(* CODESYS project listofstring.library
   DefaultNamespace: KOSTAL.TC3.Components.listOfString
   DocFormat: reStructuredText
   Description: V2019.2.1.0 - Bugfix: Delete zero pointer
      V2019.2.0.0 - now it is possible to add en empty Line.
      2019.5.0.0 - ListOfString High Performance - Add extended class ListOfString_HP with dynamic storage.
      The temporary load on the router's memory is halved.
   Author: Frank Dümpelmann
   Title: KOSTAL.TC3.Components.listOfString
   Version: 2019.5.0.0
   Company: KOSTAL GmbH & Co.KG
   Placeholder: KOSTAL.TC3.Components.listOfString

Project tree, tasks and I/O mapping:
  libraries: KOSTAL.TC3.Core.functionResponse, 2019.1.0.0 (KOSTAL GmbH & Co.KG); KOSTAL.TC3.Core.Settings, 2019.0.1.0 (KOSTAL GmbH & Co.KG); KOSTAL.TC3.Core.System, 2019.0.0.0 (KOSTAL GmbH & Co.KG); Tc2_Standard, 3.3.3.0 (Beckhoff Automation GmbH); Tc2_System, 3.5.3.0 (Beckhoff Automation GmbH); Tc2_Utilities, 3.3.54.0 (Beckhoff Automation GmbH)
  listOfString_255/
    function block FB_ListOfString_255 [ST]: _stackGetSize, addLine, clear, FB_exit, FB_init, line_GET, line_SET, maxLine, numberOfLines_GET, removeLine
    interface I_ListOfString_255: line_GET, maxLine, numberOfLines_GET
    interface I_ListOfString_255_Owner: addLine, clear, line_GET, line_SET, maxLine, numberOfLines_GET, removeLine
  ListOfString_HP/
    0_Core/
      BaseElement/
        data type P_List
        data type ST_List
      function block FB_Core [ST]: _addItem, _findItem, _findItemByIndex, _insertItem, _removeFromBegin, _removeFromEnd, _removeItem, _removeItemByIndex, _nextItem, _previousItem, _clearResult, _setResultFail, _setResultPass, _checkConsistency, _clear, _NumberOfMember, FB_exit, FB_init
      interface I_Core
      interface I_Core_Owner
    1_Base/
      function block FB_Base [ST]: _FIFO_peek, _FIFO_pop, _FIFO_push, _addMember, _findMember, _findMemberByIndex, _insertMember, _removeFromBegin, _removeFromEnd, _removeMember, _removeMemberByIndex, _clear, FB_exit, FB_init
      interface I_Base
      interface I_Base_Owner
    function block FB_ListOfString_HP [ST]: addLine, clear, line_GET, line_SET, maxLine, maxLine_udi, NumberOfLines, numberOfLines_GET, removeLine
    interface I_ListOfString_HP: maxLine_udi, NumberOfLines
    interface I_ListOfString_HP_Owner: maxLine_udi, NumberOfLines
  Project Information/
    function F_GetCompany [ST]
    function F_GetTitle [ST]
    function F_GetVersion [ST]
  Version/
    global variables Global_Version
*)

// ListOfString_HP/0_Core/BaseElement/P_List
//Pointer to an element of List
TYPE P_List : POINTER TO ST_List; END_TYPE

// ListOfString_HP/0_Core/BaseElement/ST_List
{attribute 'enable_dynamic_creation'}
TYPE ST_List :
	STRUCT
			pNext	 		: P_List;				//Pointer to next Item
			Member			: KOSTAL_TC3_Core_Settings.T_MaxString;	//Text content
			pPrevious : P_List;				//Pointer to previous item
	END_STRUCT
END_TYPE

// Version/Global_Version
{attribute 'TcGenerated'}
{attribute 'no-analysis'}
{attribute 'linkalways'}
// This function has been automatically generated from the project information.
VAR_GLOBAL CONSTANT
	{attribute 'const_non_replaced'}
	stLibVersion_KOSTAL_TC3_Components_listOfString : ST_LibVersion := (iMajor := 2019, iMinor := 5, iBuild := 0, iRevision := 0, nFlags := 1, sVersion := '2019.5.0.0');
END_VAR

// listOfString_255/FB_ListOfString_255
{attribute 'obsolete' := 'Use instead FB_ListOfString_HP'} 
(*

:Author: Frank Dümpelmann <f.duempelmann@kostal.com>, Martin Hundt <m.hundt@kostal.com>
:Date: 2018-11-19

Function
========
Keeps a list of string(255) with a variable number of elements

Usage notes
===============
| Call Method addLine to add a string at the end of the list 
| Call Method getLine to read a string from the list
| numberOfLines_GET returns the actual numer of elements in the list
| List indices are 1-based
| Suitable to implement LIFO or FIFO stacks (see example in fileLogger)

Methods and Properties
======================
| See bottom of this document for a detailed description of each method or property
| Methods starting with an underline(_) are internally used and can be ignored by the user

Usage sample:
=============

.. code:: 

	PROGRAM MAIN
	VAR
		_list	: FB_ListOfString_255;
		_i		: UINT;
		_listContent : ARRAY [1..10] OF STRING(255);
		_filled :BOOL;
	END_VAR
	
	IF NOT _filled THEN	//Add lines to the list ONCE
		_list.addLine('Line 1');
		_list.addLine('Line 2');
		_list.addLine('Line 3');
		_list.addLine('Line 4');
		_list.addLine('Line 5');
		_list.addLine('Line 6');
		_list.removeLine(5);	//Delete line no. 5
		_filled := TRUE;
	END_IF
	
	//Retrieve the lines from the list
	FOR _i:=1 TO _list.numberOfLines_GET() DO
		_listContent[_i] := _list.line_GET(_i);
	END_FOR

*)
FUNCTION_BLOCK PUBLIC FB_ListOfString_255 IMPLEMENTS I_ListOfString_255, I_ListOfString_255_Owner
VAR_INPUT
END_VAR
VAR_OUTPUT
END_VAR

VAR
	_pStack			: POINTER TO KOSTAL_TC3_Core_Settings.T_MaxString;
	_pNewStack	: POINTER TO KOSTAL_TC3_Core_Settings.T_MaxString;
	_line				:	KOSTAL_TC3_Core_Settings.T_MaxString;

	_elements	: UINT;
	_sizeLine	: UDINT;

	_maxLine	:	UINT:= 100;
END_VAR

METHOD PROTECTED _stackGetSize :	UDINT
VAR_INPUT
END_VAR

IF _pStack = 0 THEN
	_stackGetSize:= 0;
ELSE
	_stackGetSize:= SIZEOF(_line) * _elements;
END_IF
END_METHOD

(*
Description
===========
| Adds a line to end of the list
| Parameters:
| 	line: STRING(255): Text to add to the list
| Returns false in case line is empty or list is full
*)

METHOD PUBLIC addLine : BOOL
VAR_INPUT
	newLine	: KOSTAL_TC3_Core_Settings.T_MaxString;
END_VAR

VAR
	_newNumberOfElements	: UINT;
END_VAR

addLine:= FALSE;

//IF newLine = '' THEN RETURN;	END_IF
IF _elements >= _maxLine THEN RETURN;	END_IF

_newNumberOfElements	:= _elements + 1;

_pNewStack:= __NEW(STRING(255), _newNumberOfElements);

IF _elements > 0 THEN
	MEMCPY(destAddr:= ADR(_pNewStack[0]), srcAddr:= ADR(_pStack[0]), n:= _stackGetSize());
END_IF

_pNewStack[_newNumberOfElements - 1]:= newLine;

IF (_pStack <> 0) THEN	__DELETE(_pStack);	END_IF
_elements:= _newNumberOfElements;
_pStack:= __NEW(STRING(255), _elements);

MEMCPY(destAddr:= ADR(_pStack[0]), srcAddr:= ADR(_pNewStack[0]), n:= _stackGetSize());
IF (_pNewStack <> 0) THEN __DELETE(_pNewStack); END_IF

addLine:= TRUE;
END_METHOD

(*
Description
===========
| Clears the list's contents
*)
METHOD PUBLIC clear
VAR_INPUT
END_VAR

IF (_pStack <> 0) THEN __DELETE(_pStack); END_IF
IF (_pNewStack <> 0) THEN __DELETE(_pNewStack); END_IF

_elements:= 0;
END_METHOD

(*
Description
===========
| This method is called automatically
| Do not call manually 
*)
METHOD FB_exit : BOOL
VAR_INPUT
	bInCopyCode : BOOL; // if TRUE, the exit method is called for exiting an instance that is copied afterwards (online change).
END_VAR

IF (_pStack <> 0) THEN __DELETE(_pStack);	END_IF
IF (_pNewStack <> 0) THEN __DELETE(_pNewStack);	END_IF

_elements:= 0;
END_METHOD

(*
Description
===========
| This method is called automatically
| Do not call manually 
*)
METHOD FB_init : BOOL
VAR_INPUT
	bInitRetains : BOOL; // if TRUE, the retain variables are initialized (warm start / cold start)
	bInCopyCode : BOOL;  // if TRUE, the instance afterwards gets moved into the copy code (online change)
END_VAR

IF (_pStack <> 0) THEN __DELETE(_pStack);	END_IF
IF (_pNewStack <> 0) THEN __DELETE(_pNewStack);	END_IF

_elements:= 0;
END_METHOD

(*
Description
===========
| Returns the line at the given index
| Parameters:
| 	numberOfLine: index
*)
METHOD PUBLIC line_GET : KOSTAL_TC3_Core_Settings.T_MaxString
VAR_INPUT
	numberOfLine	:	UINT;	//1..numberOfLines_GET()
END_VAR

line_GET:= '';

IF numberOfLine = 0	THEN	RETURN;	END_IF
IF numberOfLine > _elements THEN	RETURN;	END_IF

line_GET	:=	_pStack[numberOfLine - 1];
END_METHOD

(*
Description
===========
| Returns the line at the given index
| Parameters:
| 	numberOfLine: index
*)
METHOD PUBLIC line_SET : BOOL
VAR_INPUT
	line	: KOSTAL_TC3_Core_Settings.T_MaxString;
	numberOfLine	:	UINT;	//1..numberOfLines_GET()
END_VAR

line_SET:= FALSE;

IF numberOfLine = 0	THEN	RETURN;	END_IF
IF numberOfLine > _elements THEN	RETURN;	END_IF

_pStack[numberOfLine - 1]:= line;

line_SET:= TRUE;
END_METHOD

(*
Description
===========
| **Maximum** number of elements in the list. 
| If the list is full, added lines will be ignored
*)
PROPERTY PUBLIC maxLine : UINT
GET

maxLine:= _maxLine;
END_GET
SET

_maxLine:= maxLine;
END_SET
END_PROPERTY

(*
Description
===========
| Returns the **actual** number of elements in the list
*)
METHOD PUBLIC numberOfLines_GET : UINT
VAR_INPUT
END_VAR

numberOfLines_GET:= _elements;
END_METHOD

(*
Description
===========
| Remove the line with the given index
| Elements after the index move up one position
| Parameters:
| 	index: line to remove
*)

METHOD PUBLIC removeLine
VAR_INPUT
	numberOfLine	:	UINT;	//1..numberOfLines_GET()
END_VAR

VAR
	_indexOfLine		: UINT;
END_VAR


IF numberOfLine = 0 THEN	RETURN;	END_IF
IF numberOfLine > _elements THEN	RETURN;	END_IF

_indexOfLine:= numberOfLine - 1;

_pStack[_indexOfLine]	:= '';

_pNewStack	:=	__NEW(STRING(255), (_elements - 1));

//if not first entry
IF _indexOfLine > 0 THEN
	MEMCPY(destAddr:= ADR(_pNewStack[0]), srcAddr:= ADR(_pStack[0]), n:= SIZEOF(_line) * _indexOfLine);
END_IF

//if not last entry
IF _indexOfLine < _elements - 1 THEN
	MEMCPY(destAddr:= ADR(_pNewStack[_indexOfLine]), srcAddr:= ADR(_pStack[numberOfLine]), n:= SIZEOF(_line) * (_elements - numberOfLine));
END_IF


IF (_pStack <> 0) THEN __DELETE(_pStack);	END_IF

_elements:= _elements - 1;
_pStack:= __NEW(STRING(255), _elements);

MEMCPY(destAddr:= ADR(_pStack[0]), srcAddr:= ADR(_pNewStack[0]), n:= _stackGetSize());
IF (_pNewStack <> 0) THEN __DELETE(_pNewStack);	END_IF
END_METHOD

END_FUNCTION_BLOCK

// ListOfString_HP/FB_ListOfString_HP
(*
	List of String
	HP -High Performance
	The temporary load on the router's memory is halved.
*)
FUNCTION_BLOCK PUBLIC FB_ListOfString_HP EXTENDS FB_Base IMPLEMENTS I_ListOfString_HP, I_ListOfString_HP_Owner
VAR
	_maxLine	: UDINT:= UDINT#16#FFFF_FFFF;
END_VAR

(*
Description
===========
| Adds a line to end of the list
| Parameters:
| 	line: STRING(255): Text to add to the list
| Returns false in case line is empty or list is full
*)
METHOD addLine : BOOL
VAR_INPUT
	newLine	: KOSTAL_TC3_Core_Settings.T_MaxString;
END_VAR

VAR
	_fRes: KOSTAL_TC3_Core_functionResponse.FB_functionResponse;
END_VAR

addLine:= SUPER^._addMember(newLine, _fRes) AND _fRes.success;
END_METHOD

(*
Description
===========
| Clears the list's contents
*)
METHOD clear

SUPER^._clear();
END_METHOD

(*
Description
===========
| Returns the line at the given index
| Parameters:
| 	numberOfLine: index
*)
METHOD line_GET : KOSTAL_TC3_Core_Settings.T_MaxString
VAR_INPUT
	(*1..numberOfLines_GET()*)
	numberOfLine	: UINT;
END_VAR

VAR
	_fRes: KOSTAL_TC3_Core_functionResponse.FB_functionResponse;
END_VAR

_findMemberByIndex(NumberOfLine - 1, line_GET, _fRes);
END_METHOD

(*
Description
===========
| Returns the line at the given index
| Parameters:
| 	numberOfLine: index
*)
METHOD line_SET : BOOL
VAR_INPUT
	line	: KOSTAL_TC3_Core_Settings.T_MaxString;
	(*1..numberOfLines_GET()*)
	numberOfLine	: UINT;
END_VAR

VAR
	_item: P_List;
	_fRes: KOSTAL_TC3_Core_functionResponse.FB_functionResponse;
END_VAR

IF NOT SUPER^._findItemByIndex(numberOfLine - 1, _item, _fRes)	THEN RETURN;	END_IF

IF NOT _fRes.success	THEN RETURN;	END_IF

IF _item = 0 THEN RETURN;	END_IF

_item^.Member:= line;

line_SET:= TRUE;
END_METHOD

(*
Description
===========
| **Maximum** number of elements in the list. 
| If the list is full, added lines will be ignored
*)
PROPERTY maxLine : UINT
GET

IF _maxLine	> UDINT#16#0000_FFFF THEN	maxLine:= UINT#16#FFFF;
ELSE																	maxLine:= UDINT_TO_UINT(_maxLine);
END_IF
END_GET
SET

_maxLine:= UINT_TO_UDINT(maxLine);
END_SET
END_PROPERTY

(*
Description
===========
| **Maximum** number of elements in the list. 
| If the list is full, added lines will be ignored
*)
PROPERTY maxLine_udi : UDINT
GET

maxLine_udi:= _maxLine;
END_GET
SET

_maxLine:= maxLine_udi;
END_SET
END_PROPERTY

PROPERTY PUBLIC NumberOfLines : UDINT
GET

NumberOfLines:= SUPER^._Count;
END_GET
END_PROPERTY


(*
Description
===========
| Returns the **actual** number of elements in the list
*)
METHOD numberOfLines_GET : UINT

IF SUPER^._NumberOfMember > UDINT#16#FFFF THEN	numberOfLines_GET:= UINT#16#FFFF;
ELSE																						numberOfLines_GET:= UDINT_TO_UINT(SUPER^._NumberOfMember);
END_IF
END_METHOD

(*
Description
===========
| Remove the line with the given index
| Elements after the index move up one position
| Parameters:
| 	index: line to remove
*)
METHOD removeLine
VAR_INPUT
	(*1..numberOfLines_GET()*)
	numberOfLine	: UINT;
END_VAR

VAR
	_fRes: KOSTAL_TC3_Core_functionResponse.FB_functionResponse;
END_VAR

SUPER^._removeMemberByIndex(numberOfLine - 1, _fRes);
END_METHOD

END_FUNCTION_BLOCK

// ListOfString_HP/1_Base/FB_Base
(*

| =========================================================================
| List of Items from base Interface {KOSTAL_TC3_Core_System.I_Interface} 
| =========================================================================

..code::

	//In addition to the interface, each item contains the pointer to the previous item 
	//as well as the pointer to the next item in the list.

	TYPE ST_List :
		STRUCT
				pNext			: P_List;
				Line			: KOSTAL_TC3_Core_Settings.T_MaxString;	//Text content
				pPrevious : P_List;
		END_STRUCT
	END_TYPE

============= ======================================= ======================
| The List is defined by (p)Begin and (p)End and also the count of Members 
----------------------------------------------------------------------------
============= ======================================= ======================
 **_pBegin**  >>>>>>>>>>>>>>>>>>>>>>>>>>>>>>>>>>>>>>  **_pEnd**                     
 **Item-1**	    Item-2   Item-3   Item-4  Item-5      **Item-n**                   
============= ======================================= ======================



| =========================================================================
| The Member is an Interface as payload and an access pointer to the        
| previous member and the next member                                      
| ---------------------------------------------------------------------------
| Previous Item ---<<<Pointer-Previous-[Item]-Pointer-Next>>>---NextItem---
| =========================================================================

*)
FUNCTION_BLOCK ABSTRACT FB_Base EXTENDS FB_Core IMPLEMENTS I_Base, I_Base_Owner

VAR
END_VAR

//methode return the Member from begin 
METHOD PROTECTED _FIFO_peek : BOOL
VAR_INPUT
	FoundMember	: REFERENCE TO KOSTAL_TC3_Core_Settings.T_MaxString;	//return value
	Result			: REFERENCE TO KOSTAL_TC3_Core_functionResponse.FB_functionResponse;
END_VAR

_clearResult(Result);

IF 		NOT __ISVALIDREF(FoundMember) THEN _setResultFail(Result, 'FoundMember has no valid reference'); 
ELSE	_FIFO_peek:= _findMemberByIndex(0, FoundMember, Result);
END_IF
END_METHOD

//methode return the Member from begin and remove it from List
METHOD PROTECTED _FIFO_pop : BOOL
VAR_INPUT
	FoundMember	: REFERENCE TO KOSTAL_TC3_Core_Settings.T_MaxString;	//return value
	Result			: REFERENCE TO KOSTAL_TC3_Core_functionResponse.FB_functionResponse;
END_VAR


_clearResult(Result);

_FIFO_pop:= _findMemberByIndex(0, FoundMember, Result);

IF _FIFO_pop THEN	_FIFO_pop:= _removeFromBegin(Result);	END_IF
END_METHOD

//push/add the {Member} to begin from List
METHOD PROTECTED _FIFO_push : BOOL
VAR_INPUT
	Member	: KOSTAL_TC3_Core_Settings.T_MaxString;
	Result	: REFERENCE TO KOSTAL_TC3_Core_functionResponse.FB_functionResponse;
END_VAR


_FIFO_push:= _insertItem(UDINT#0, Member, Result);
END_METHOD

(*
	add new Member to end of list
*)
METHOD PROTECTED _addMember : BOOL

VAR_INPUT
	Member		: KOSTAL_TC3_Core_Settings.T_MaxString;
	Result	: REFERENCE TO KOSTAL_TC3_Core_functionResponse.FB_functionResponse;
END_VAR


VAR
	_Member: KOSTAL_TC3_Core_System.I_Interface;
END_VAR

_addMember:= _addItem(Member, Result);
END_METHOD

(*
	Search for the element {Item} in the list and return {FoundItem} if it is found {_findItem = TRUE}
*)
METHOD PROTECTED _findMember : BOOL
VAR_INPUT
	Member			: KOSTAL_TC3_Core_Settings.T_MaxString;
	FoundMember	: REFERENCE TO KOSTAL_TC3_Core_Settings.T_MaxString;	//return value
	Result			: REFERENCE TO KOSTAL_TC3_Core_functionResponse.FB_functionResponse;
END_VAR

VAR
	_Item		: P_List;
END_VAR

_clearResult(Result);

IF NOT __ISVALIDREF(FoundMember)			THEN _setResultFail(Result, 'FoundItem has no valid reference');	RETURN;	END_IF

_findMember:= _findItem(Member, _Item, Result);

IF NOT _findMember		THEN	RETURN;	END_IF
IF _Item = 0 					THEN	RETURN;	END_IF

FoundMember:= _Item^.Member;
END_METHOD

//find a modul by index  
METHOD PROTECTED _findMemberByIndex : BOOL
VAR_INPUT
	Index				: UDINT;	//index of item
	FoundMember	: REFERENCE TO KOSTAL_TC3_Core_Settings.T_MaxString;	//return value
	Result			: REFERENCE TO KOSTAL_TC3_Core_functionResponse.FB_functionResponse;	//result information
END_VAR

VAR
	_FoundItem	: P_List;
END_VAR

IF NOT __ISVALIDREF(FoundMember)	THEN _setResultFail(Result, 'FoundMember has no valid reference');	RETURN;	END_IF

FoundMember:= '';

_findMemberByIndex:= _findItemByIndex(Index,_FoundItem, Result);

IF NOT _findMemberByIndex THEN RETURN;	END_IF
IF _FoundItem = 0 THEN RETURN;	END_IF

FoundMember:= _FoundItem^.Member;

_findMemberByIndex:= TRUE;
END_METHOD

METHOD PROTECTED _insertMember : BOOL
VAR_INPUT
	Index		: UDINT;	//Index a which shall inserted the {Item}
	Member	: KOSTAL_TC3_Core_Settings.T_MaxString;
	Result	: REFERENCE TO KOSTAL_TC3_Core_functionResponse.FB_functionResponse;
END_VAR

VAR
	_Member: KOSTAL_TC3_Core_System.I_Interface;
END_VAR

_insertMember:= _insertItem(Index, Member, Result);
END_METHOD

(*
	remove Item from begin of list
*)
METHOD PROTECTED _removeFromBegin : BOOL
VAR_INPUT
	Result	: REFERENCE TO KOSTAL_TC3_Core_functionResponse.FB_functionResponse;
END_VAR

_removeFromBegin:= THIS^._removeMemberByIndex(0, Result);
END_METHOD

(*
	remove Item from end of list
*)
METHOD PROTECTED _removeFromEnd : BOOL
VAR_INPUT
	Result	: REFERENCE TO KOSTAL_TC3_Core_functionResponse.FB_functionResponse;
END_VAR

_removeFromEnd:= THIS^._removeMemberByIndex(_Count, Result);
END_METHOD

(*
	remove given {Member} from List
*)
METHOD PROTECTED _removeMember : BOOL
VAR_INPUT
	Member	: KOSTAL_TC3_Core_Settings.T_MaxString;
	Result	: REFERENCE TO KOSTAL_TC3_Core_functionResponse.FB_functionResponse;
END_VAR

VAR
	_Item		: P_List;
	_bFound: BOOL;
END_VAR


_bFound:= _findItem(Member, _Item, Result);

IF NOT _bFound THEN RETURN;	END_IF

_removeMember:= _removeItem(_Item, Result);
END_METHOD

(*
	remove given {Index} from List
*)
METHOD PROTECTED _removeMemberByIndex : BOOL
VAR_INPUT
	Index		: UDINT;
	Result	: REFERENCE TO KOSTAL_TC3_Core_functionResponse.FB_functionResponse;
END_VAR

VAR
	_bFound	: BOOL;
	_Member	: KOSTAL_TC3_Core_Settings.T_MaxString;

END_VAR

IF NOT _findMemberByIndex(Index, _Member, Result)	THEN RETURN;	END_IF

_removeMemberByIndex:= _removeMember(_Member, Result);
END_METHOD

(*
	Delete the complete content of the list
*)
METHOD PROTECTED _clear
VAR_INPUT
END_VAR

WHILE THIS^._pBegin <> 0 DO
    THIS^._removeMember(THIS^._pBegin^.Member, 0);  
END_WHILE
END_METHOD

METHOD FB_exit : BOOL
VAR_INPUT
	bInCopyCode : BOOL; // if TRUE, the exit method is called for exiting an instance that is copied afterwards (online change).
END_VAR

_clear();
END_METHOD

METHOD FB_init : BOOL
VAR_INPUT
	bInitRetains : BOOL; // if TRUE, the retain variables are initialized (warm start / cold start)
	bInCopyCode : BOOL;  // if TRUE, the instance afterwards gets moved into the copy code (online change)
END_VAR

_clear();
END_METHOD

END_FUNCTION_BLOCK

// ListOfString_HP/0_Core/FB_Core
(*

| =========================================================================
| List of Items from base Interface {KOSTAL_TC3_Core_System.I_Interface} 
| =========================================================================

..code::

	//In addition to the interface, each item contains the pointer to the previous item 
	//as well as the pointer to the next item in the list.

	TYPE ST_List :
		STRUCT
				pNext			: P_List;
				iMember		: KOSTAL_TC3_Core_System.I_Interface;	
				pPrevious : P_List;
		END_STRUCT
	END_TYPE

============= ======================================= ======================
| The List is defined by (p)Begin and (p)End and also the count of Members 
----------------------------------------------------------------------------
============= ======================================= ======================
 **_pBegin**  >>>>>>>>>>>>>>>>>>>>>>>>>>>>>>>>>>>>>>  **_pEnd**                     
 **Item-1**	    Item-2   Item-3   Item-4  Item-5      **Item-n**                   
============= ======================================= ======================



| =========================================================================
| The Member is an Interface as payload and an access pointer to the        
| previous member and the next member                                      
| ---------------------------------------------------------------------------
| Previous Item ---<<<Pointer-Previous-[Item]-Pointer-Next>>>---NextItem---
| =========================================================================

*)
FUNCTION_BLOCK ABSTRACT FB_Core IMPLEMENTS I_Core, I_Core_Owner

VAR
	_pBegin	: P_List;	//origin of List
  _pEnd		: P_List;	//end of List
	_Count	: UDINT;	//number of registered Member
END_VAR

(*
	add new item to end of list
*)
METHOD PROTECTED _addItem : BOOL

VAR_INPUT
	Member		: KOSTAL_TC3_Core_Settings.T_MaxString;
	Result	: REFERENCE TO KOSTAL_TC3_Core_functionResponse.FB_functionResponse;
END_VAR

VAR
	_pNewItem	: P_List;
END_VAR
_clearResult(Result);

//IF Item = 0 THEN _setResultFail(Result, 'Parameter Item is empty');	RETURN;	END_IF


//create a new Item
_pNewItem:= __NEW(ST_List);

//If creation failed 
IF _pNewItem = 0 THEN _setResultFail(Result, 'New Item cannot create');	RETURN;	END_IF

//If list is empty
IF THIS^._Count = 0 (*THIS^._pEnd = 0*) THEN THIS^._pBegin:= THIS^._pEnd:= _pNewItem; 
ELSE

	//set new item previous item to actual last item (THIS^._pEnd)
	_pNewItem^.pPrevious:= THIS^._pEnd;
	_pNewItem^.pPrevious^.pNext:= _pNewItem;
 
	THIS^._pEnd:= _pNewItem;
END_IF

THIS^._pEnd^.Member:= Member;
THIS^._Count:= THIS^._Count + UDINT#1;

_setResultPass(Result, 'addItem successful');

_addItem:= TRUE;
END_METHOD

(*
	Search for the element {Item} in the list and return {FoundItem} if it is found {_findItem = TRUE}
*)
METHOD PROTECTED _findItem : BOOL
VAR_INPUT
	Member		: KOSTAL_TC3_Core_Settings.T_MaxString;
	FoundItem	: REFERENCE TO P_List;
	Result		: REFERENCE TO KOSTAL_TC3_Core_functionResponse.FB_functionResponse;
END_VAR

VAR
	_Item		: P_List;
END_VAR
_clearResult(Result);

IF NOT __ISVALIDREF(FoundItem)	THEN _setResultFail(Result, 'FoundItem has no valid reference');	RETURN;	END_IF


_Item := THIS^._pBegin;

WHILE _Item <> 0 DO

	IF _Item^.Member = Member THEN

		FoundItem := _Item;

		_findItem:= TRUE;

		_setResultPass(Result, 'Item found');
		
		RETURN;   

	END_IF
	
	_Item := THIS^._nextItem(_Item, 0);

END_WHILE

//FoundItem:= _Item;

_setResultFail(Result, 'Item not found');

_findItem:= FALSE;
END_METHOD

(*
	Search for the element {Item} in the list and return {FoundItem} if it is found {_findItem = TRUE}
*)
METHOD PROTECTED _findItemByIndex : BOOL
VAR_INPUT
	Index			: UDINT;
	FoundItem	: REFERENCE TO P_List;
	Result		: REFERENCE TO KOSTAL_TC3_Core_functionResponse.FB_functionResponse;
END_VAR

VAR
	_Item		: P_List;
	_udi: UDINT;
END_VAR

_findItemByIndex:= FALSE;

_clearResult(Result);

IF _Count = 0										THEN _setResultFail(Result, 'List is empty');											RETURN;	END_IF
IF Index > (_Count - 1)					THEN _setResultFail(Result, 'Parameter Index is out of range');		RETURN;	END_IF
IF NOT __ISVALIDREF(FoundItem)	THEN _setResultFail(Result, 'FoundItem has no valid reference');	RETURN;	END_IF


_Item := THIS^._pBegin;

IF Index > 0 THEN
	FOR _udi:= 0 TO Index - 1 DO
			_Item := THIS^._nextItem(_Item, 0);
	END_FOR
END_IF

FoundItem:= _Item;

IF FoundItem = 0 THEN
	_setResultFail(Result, 'Item not found');
ELSE	
	_setResultPass(Result, 'Item found');
	_findItemByIndex:= TRUE;
END_IF
END_METHOD

METHOD PROTECTED _insertItem : BOOL
VAR_INPUT
	Index		: UDINT;	//Index a which shall inserted the {Item}
	Member	: KOSTAL_TC3_Core_Settings.T_MaxString;
	Result	: REFERENCE TO KOSTAL_TC3_Core_functionResponse.FB_functionResponse;
END_VAR

VAR
	_pNewItem			: P_List;
	_pExitingItem	: P_List;
END_VAR
_clearResult(Result);

//if List is empty add item 
IF (Index = 0) AND (_Count = 0)	THEN _insertItem:= _addItem(Member, Result);	RETURN;	END_IF

//Index is in list not available 
IF Index > (_Count - 1) THEN _setResultFail(Result, 'Index is out of range');	RETURN;	END_IF

//if index is end of list then add item to end of list 
IF (Index = (_Count - 1)) THEN _insertItem:= _addItem(Member, Result);	RETURN;	END_IF

//try to find item where shall inserted
IF NOT _findItemByIndex(Index, _pExitingItem, Result) THEN RETURN;	END_IF
IF _pExitingItem = 0 THEN _setResultFail(Result, 'Item not available');	RETURN;	END_IF


//create a new Item
_pNewItem:= __NEW(ST_List);

//If creation failed 
IF _pNewItem = 0 THEN _setResultFail(Result, 'New Item cannot create');	RETURN;	END_IF

_pNewItem^.Member:= Member;

_pNewItem^.pNext		:= _pExitingItem;							//set the next item from new item to existing founded item
_pNewItem^.pPrevious:= _pExitingItem^.pPrevious;	//set the previous from existing item to the previous of new item

//if a previous exist then
//set the next from previous from existing item to the previous of new item
IF _pNewItem^.pPrevious <> 0 THEN	_pNewItem^.pPrevious^.pNext:= _pNewItem;	END_IF

_pExitingItem^.pPrevious:= _pNewItem;							//set the previous from existing founded item to  new item

//if inserted at the begin of list, set the begin pointer to new Item
IF THIS^._pBegin = _pExitingItem THEN	THIS^._pBegin:= _pNewItem;	END_IF

THIS^._Count:= THIS^._Count + UDINT#1;

_setResultPass(Result, 'insertItem successful');

_insertItem:= TRUE;
END_METHOD

(*
	remove Item from begin of list
*)
METHOD PROTECTED _removeFromBegin : BOOL
VAR_INPUT
	Result	: REFERENCE TO KOSTAL_TC3_Core_functionResponse.FB_functionResponse;
END_VAR

_removeFromBegin:= THIS^._removeItemByIndex(0, Result);
END_METHOD

(*
	remove Item from end of list
*)
METHOD PROTECTED _removeFromEnd : BOOL
VAR_INPUT
	Result	: REFERENCE TO KOSTAL_TC3_Core_functionResponse.FB_functionResponse;
END_VAR

_removeFromEnd:= THIS^._removeItemByIndex(_Count, Result);
END_METHOD

(*
	remove given {Item} from List
*)
METHOD PROTECTED _removeItem : BOOL
VAR_INPUT
	Item		: P_List;
	Result	: REFERENCE TO KOSTAL_TC3_Core_functionResponse.FB_functionResponse;
END_VAR

_clearResult(Result);

IF Item = 0 THEN _setResultFail(Result, 'Parameter Item is empty');	RETURN;	END_IF

//exist a next member
IF Item^.pNext <> 0 THEN
	//set next members previous Item  to my previous Item
	Item^.pNext^.pPrevious := Item^.pPrevious; 
END_IF

//exist a previous member
IF Item^.pPrevious <> 0 THEN
	//set previous members next Item  to my next Item
	Item^.pPrevious^.pNext := Item^.pNext;
END_IF

//Item is the once member
IF Item = THIS^._pBegin AND Item = THIS^._pEnd THEN
	
	THIS^._pBegin := 0;
	THIS^._pEnd := 0;

ELSIF Item = THIS^._pBegin (*AND Item <> THIS^._pEnd*) THEN

	THIS^._pBegin := Item^.pNext;

ELSIF (*Item <> THIS^._pBegin AND*) Item = THIS^._pEnd THEN

	THIS^._pEnd := Item^.pPrevious;

END_IF

__DELETE(Item);

IF  THIS^._Count > UDINT#0 THEN	THIS^._Count := THIS^._Count - UDINT#1;	
ELSE
	_setResultFail(Result, 'removeItem Counter underflow');
	RETURN;
END_IF

_setResultPass(Result, 'removeItem successful');
_removeItem:= TRUE;
END_METHOD

(*
	remove given {Index} from List
*)
METHOD PROTECTED _removeItemByIndex : BOOL
VAR_INPUT
	Index		: UDINT;
	Result	: REFERENCE TO KOSTAL_TC3_Core_functionResponse.FB_functionResponse;
END_VAR

VAR
	_Item		: P_List;
	_bFound	: BOOL;
END_VAR

IF NOT _findItemByIndex(Index, _Item, Result)	THEN RETURN;	END_IF

_removeItemByIndex:= _removeItem(_Item, Result);
END_METHOD

// retreives the pointer to the next item of the given entry
METHOD PROTECTED _nextItem : P_List;
VAR_INPUT
    Item : P_List;
		Result	: REFERENCE TO KOSTAL_TC3_Core_functionResponse.FB_functionResponse;
END_VAR
VAR
	_Res	: P_List;
END_VAR

IF Item <> 0 THEN	_Res := Item^.pNext;
ELSE							_Res := 0;
END_IF

_nextItem:= _Res;
END_METHOD

// retreives the previous item of the given entry
METHOD PROTECTED _previousItem : P_List
VAR_INPUT
    Item 	: P_List;
END_VAR
VAR
	_Res	: P_List;
END_VAR

IF Item <> 0 THEN	_Res := Item^.pPrevious;
ELSE							_Res := 0;
END_IF

_previousItem:= _Res;
END_METHOD

(*
	Clear result component
*)
METHOD PROTECTED _clearResult : BOOL
VAR_INPUT
	IN : REFERENCE TO KOSTAL_TC3_Core_functionResponse.FB_functionResponse;
END_VAR

IF __ISVALIDREF(IN) THEN IN.clear(); _clearResult:= TRUE;	END_IF
END_METHOD

(*
	set result to fail with given information 
*)
METHOD PROTECTED _setResultFail : BOOL
VAR_INPUT
	IN : REFERENCE TO KOSTAL_TC3_Core_functionResponse.FB_functionResponse;
	Info	: KOSTAL_TC3_Core_Settings.T_MaxString;
END_VAR

IF __ISVALIDREF(IN) THEN 

	IN.success:= FALSE;
	IN.status:= Info;

	_setResultFail:= TRUE;

END_IF
END_METHOD

(*
	set result to pass with given information 
*)
METHOD PROTECTED _setResultPass : BOOL
VAR_INPUT
	IN : REFERENCE TO KOSTAL_TC3_Core_functionResponse.FB_functionResponse;
	Info	: KOSTAL_TC3_Core_Settings.T_MaxString;
END_VAR

IF __ISVALIDREF(IN) THEN 

	IN.success:= TRUE;
	IN.status:= Info;

	_setResultPass:= TRUE;

END_IF
END_METHOD

(*
	Check if the list is consistent
*)
METHOD PROTECTED _checkConsistency : BOOL
VAR_INPUT
	Result	: REFERENCE TO KOSTAL_TC3_Core_functionResponse.FB_functionResponse;
END_VAR

VAR
	_pItem			: P_List;
	_pNext			: P_List;
	_pPrev			: P_List;
	_nItemCounter	: UDINT;
	_bBeginOk			: BOOL;
	_bEndOk			: BOOL;
	_bPrevLinkOk		: BOOL;
	_bNextLinkOk		: BOOL;
	_bItemCountOk	: BOOL;
END_VAR
// check from pHead to pTail
_pItem:= THIS^._pBegin;
_nItemCounter:= 0;

IF THIS^._pBegin <> 0 THEN
	_bBeginOk:= (THIS^._pBegin^.pPrevious = 0);
ELSE
	_bBeginOk:= TRUE;
END_IF

IF THIS^._pEnd <> 0 THEN
	_bEndOk:= (THIS^._pEnd^.pNext = 0);
ELSE
	_bEndOk:= TRUE;
END_IF

IF _bBeginOk AND _bEndOk THEN

	_bPrevLinkOk:= TRUE;
	_bNextLinkOk:= TRUE;

	WHILE _pItem <> 0 DO
		
		_pPrev:= _pItem^.pPrevious;
		_pNext:= _pItem^.pNext;

		IF _pPrev <> 0 THEN
			_bPrevLinkOk:= (_pPrev^.pNext = _pItem);
		ELSE
			_bPrevLinkOk:= (_pItem = THIS^._pBegin);
		END_IF

		IF _pNext <> 0 THEN
			_bNextLinkOk:= (_pNext^.pPrevious = _pItem);
		ELSE
			_bNextLinkOk:= (_pItem = THIS^._pEnd);
		END_IF

		IF NOT _bNextLinkOk OR NOT _bPrevLinkOk THEN	EXIT;	END_IF

		//handle iteration
		_nItemCounter:= _nItemCounter + UDINT#1;
		_pItem:= THIS^._nextItem(_pItem, 0);

	END_WHILE

END_IF

_bItemCountOk:= (_nItemCounter = THIS^._Count);

IF 		NOT _bBeginOk			THEN	_setResultFail(Result, 'List head not ok');
ELSIF NOT _bEndOk				THEN	_setResultFail(Result, 'List End not ok');
ELSIF NOT _bPrevLinkOk 	THEN	_setResultFail(Result, Tc2_Standard.CONCAT('Previous Link failed by item ', UDINT_TO_STRING(_nItemCounter)));
ELSIF NOT _bNextLinkOk	THEN	_setResultFail(Result, Tc2_Standard.CONCAT('Next Link failed by item ', UDINT_TO_STRING(_nItemCounter)));
ELSIF NOT	_bItemCountOk THEN	_setResultFail(Result, 'Itemcounter is not ok');
ELSE													_setResultPass(Result, 'List is consistent');	_checkConsistency:= TRUE;
END_IF
END_METHOD

(*
	Delete the complete content of the list
*)
METHOD PROTECTED _clear

WHILE THIS^._pBegin <> 0 DO
    THIS^._removeItem(THIS^._pBegin, 0);  
END_WHILE
END_METHOD

//return the nnumber of items in List
PROPERTY PROTECTED _NumberOfMember : UDINT
GET

_NumberOfMember:= _Count;
END_GET
END_PROPERTY

METHOD FB_exit : BOOL
VAR_INPUT
	bInCopyCode : BOOL; // if TRUE, the exit method is called for exiting an instance that is copied afterwards (online change).
END_VAR

_clear();
END_METHOD

METHOD FB_init : BOOL
VAR_INPUT
	bInitRetains : BOOL; // if TRUE, the retain variables are initialized (warm start / cold start)
	bInCopyCode : BOOL;  // if TRUE, the instance afterwards gets moved into the copy code (online change)
END_VAR

_clear();
END_METHOD

END_FUNCTION_BLOCK

// ListOfString_HP/0_Core/I_Core
INTERFACE I_Core EXTENDS KOSTAL_TC3_Core_System.I_Interface

END_INTERFACE

// ListOfString_HP/0_Core/I_Core_Owner
INTERFACE I_Core_Owner EXTENDS KOSTAL_TC3_Core_System.I_Interface

END_INTERFACE

// ListOfString_HP/1_Base/I_Base
INTERFACE I_Base EXTENDS I_Core

END_INTERFACE

// ListOfString_HP/1_Base/I_Base_Owner
INTERFACE I_Base_Owner EXTENDS I_Core_Owner

END_INTERFACE

// ListOfString_HP/I_ListOfString_HP
INTERFACE I_ListOfString_HP EXTENDS I_ListOfString_255

(*
Description
===========
| **Maximum** number of elements in the list. 
| If the list is full, added lines will be ignored
*)
PROPERTY maxLine_udi : UDINT
GET
END_GET
END_PROPERTY

PROPERTY PUBLIC NumberOfLines : UDINT
GET
END_GET
END_PROPERTY

END_INTERFACE

// listOfString_255/I_ListOfString_255
INTERFACE I_ListOfString_255 EXTENDS KOSTAL_TC3_Core_System.I_Interface

(*
Description
===========
| Returns the line at the given index
| Parameters:
| 	numberOfLine: index
*)
METHOD PUBLIC line_GET : KOSTAL_TC3_Core_Settings.T_MaxString
VAR_INPUT
	numberOfLine	:	UINT;	//1..numberOfLines_GET()
END_VAR
END_METHOD

(*
Description
===========
| **Maximum** number of elements in the list. 
| If the list is full, added lines will be ignored
*)
PROPERTY PUBLIC maxLine : UINT
GET
END_GET
END_PROPERTY

(*
Description
===========
| Returns the **actual** number of elements in the list
*)
METHOD PUBLIC numberOfLines_GET : UINT
VAR_INPUT
END_VAR
END_METHOD

END_INTERFACE

// ListOfString_HP/I_ListOfString_HP_Owner
INTERFACE I_ListOfString_HP_Owner EXTENDS I_ListOfString_255_Owner

(*
Description
===========
| **Maximum** number of elements in the list. 
| If the list is full, added lines will be ignored
*)
PROPERTY maxLine_udi : UDINT
GET
END_GET
SET
END_SET
END_PROPERTY

PROPERTY PUBLIC NumberOfLines : UDINT
GET
END_GET
END_PROPERTY

END_INTERFACE

// listOfString_255/I_ListOfString_255_Owner
INTERFACE I_ListOfString_255_Owner EXTENDS KOSTAL_TC3_Core_System.I_Interface

(*
Description
===========
| Adds a line to end of the list
| Parameters:
| 	line: STRING(255): Text to add to the list
| Returns false in case line is empty or list is full
*)

METHOD PUBLIC addLine : BOOL
VAR_INPUT
	newLine	: KOSTAL_TC3_Core_Settings.T_MaxString;
END_VAR
END_METHOD

(*
Description
===========
| Clears the list's contents
*)
METHOD PUBLIC clear
VAR_INPUT
END_VAR
END_METHOD

(*
Description
===========
| Returns the line at the given index
| Parameters:
| 	numberOfLine: index
*)
METHOD PUBLIC line_GET : KOSTAL_TC3_Core_Settings.T_MaxString
VAR_INPUT
	numberOfLine	:	UINT;	//1..numberOfLines_GET()
END_VAR
END_METHOD

(*
Description
===========
| Returns the line at the given index
| Parameters:
| 	numberOfLine: index
*)
METHOD PUBLIC line_SET : BOOL
VAR_INPUT
	line	: KOSTAL_TC3_Core_Settings.T_MaxString;
	numberOfLine	:	UINT;	//1..numberOfLines_GET()
END_VAR
END_METHOD

(*
Description
===========
| **Maximum** number of elements in the list. 
| If the list is full, added lines will be ignored
*)
PROPERTY PUBLIC maxLine : UINT
GET
END_GET
SET
END_SET
END_PROPERTY

(*
Description
===========
| Returns the **actual** number of elements in the list
*)
METHOD PUBLIC numberOfLines_GET : UINT
VAR_INPUT
END_VAR
END_METHOD

(*
Description
===========
| Remove the line with the given index
| Elements after the index move up one position
| Parameters:
| 	index: line to remove
*)

METHOD PUBLIC removeLine
VAR_INPUT
	numberOfLine	:	UINT;	//1..numberOfLines_GET()
END_VAR
END_METHOD

END_INTERFACE

// Project Information/F_GetCompany
// This function has been automatically generated from the project information.
{attribute 'signature_flag' := '1073741824'}
{attribute 'TcGenerated'}
{attribute 'no-analysis'}
FUNCTION F_GetCompany : WSTRING
VAR_INPUT
	
END_VAR

F_GetCompany := "KOSTAL GmbH & Co.KG";

END_FUNCTION

// Project Information/F_GetTitle
// This function has been automatically generated from the project information.
{attribute 'signature_flag' := '1073741824'}
{attribute 'TcGenerated'}
{attribute 'no-analysis'}
FUNCTION F_GetTitle : WSTRING
VAR_INPUT
	
END_VAR

F_GetTitle := "KOSTAL.TC3.Components.listOfString";

END_FUNCTION

// Project Information/F_GetVersion
// This function has been automatically generated from the project information.
{attribute 'signature_flag' := '1073741824'}
{attribute 'TcGenerated'}
{attribute 'no-analysis'}
FUNCTION F_GetVersion : ST_LibVersion
VAR_INPUT
	
END_VAR

F_GetVersion.iMajor := 2019;
F_GetVersion.iMinor := 5;
F_GetVersion.iBuild := 0;
F_GetVersion.iRevision := 0;
F_GetVersion.sVersion := '2019.5.0.0';
F_GetVersion.nFlags := 1;

END_FUNCTION
